Fanuc KAREL source: KA00006.KL

PROGRAM KA00006
%NOLOCKGROUP
VAR
  SRC: INTEGER
  DST: XYZWPR
BEGIN
  SRC = 2
  DST = SRC
END KA00006
